// TIA Portal V20 export
Screen "PN_DIAGNOSTIC ETH P9P10"  1276x673
  ScreenItem "Line_Header_X0_Y64" at 0,64 size 1276x0  Type=HmiLine
  ScreenItem "Title_ScreenOverview_X390_Y2" at 390,2 size 500x30  Type=HmiTextBox
  ScreenItem "PN-Diag_Reset" at 93,2 size 90x60  Type=HmiButton
  ScreenItem "PN-Diag_ReadNew" at 184,2 size 90x60  Type=HmiButton
  ScreenItem "Textfeld_1" at 292,8 size 95x22  Type=HmiTextBox
  ScreenItem "LED_1_Left_2" at 0,0 size 100x30  Type=HmiCircle
  ScreenItem "LED_1_Left_1" at 0,0 size 100x30  Type=HmiCircle
  ScreenItem "Textfeld_4" at 292,35 size 95x22  Type=HmiTextBox
  ScreenItem "permanentareaborderrectangle" at 0,0 size 0x0  Type=HmiRectangle
  ScreenItem "Button_Back" at 2,2 size 90x60  Type=HmiButton
  ScreenItem "PN-Diag_Counters" at 1093,2 size 90x60  Type=HmiButton
  ScreenItem "PN-Diag_LegendᆉY2" at 1184,2 size 90x60  Type=HmiButton
  ScreenItem "Rectangle_1" at 51,92 size 203x123  Type=HmiRectangle
  ScreenItem "LSicar_DeviceDiag_7" at 485,101 size 170x97  Type=HmiFaceplateContainer
  ScreenItem "LSicar_DeviceDiag_2" at 292,273 size 171x97  Type=HmiFaceplateContainer
  ScreenItem "LSicar_DeviceDiag_4" at 81,101 size 170x97  Type=HmiFaceplateContainer
  ScreenItem "LSicar_DeviceDiag_11" at 293,101 size 170x105  Type=HmiFaceplateContainer
  ScreenItem "LSicar_DeviceDiag_3" at 1942,495 size 170x97  Type=HmiFaceplateContainer
  ScreenItem "LSicar_DeviceDiag_5" at 485,274 size 170x97  Type=HmiFaceplateContainer
  ScreenItem "LSicar_DeviceDiag_10" at 1604,81 size 170x97  Type=HmiFaceplateContainer
  ScreenItem "LSicar_DeviceDiag_6" at 2123,495 size 170x97  Type=HmiFaceplateContainer
  ScreenItem "LSicar_DeviceDiag_16" at 1375,728 size 170x97  Type=HmiFaceplateContainer
  ScreenItem "Faceplate container_1" at 880,104 size 170x100  Type=HmiFaceplateContainer
  ScreenItem "LSicar_DeviceDiag_13" at 2023,203 size 170x97  Type=HmiFaceplateContainer
  ScreenItem "线_4" at 190,162 size 60x0  Type=HmiLine
  ScreenItem "线_6" at 253,143 size 0x19  Type=HmiLine
  ScreenItem "线_26" at 254,142 size 129x0  Type=HmiLine
  ScreenItem "LSicar_DeviceDiag_17" at 61,269 size 170x105  Type=HmiFaceplateContainer
  ScreenItem "LSicar_DeviceDiag_18" at 680,101 size 170x97  Type=HmiFaceplateContainer
  ScreenItem "线_1" at 156,162 size 0x145  Type=HmiLine
  ScreenItem "线_3" at 363,152 size 23x0  Type=HmiLine
  ScreenItem "线_5" at 156,162 size 20x0  Type=HmiLine
  ScreenItem "线_7" at 363,153 size 0x54  Type=HmiLine
  ScreenItem "线_8" at 363,207 size 220x0  Type=HmiLine
  ScreenItem "线_9" at 583,179 size 0x27  Type=HmiLine
  ScreenItem "线_10" at 376,163 size 14x0  Type=HmiLine
  ScreenItem "线_11" at 376,163 size 0x54  Type=HmiLine
  ScreenItem "线_12" at 376,217 size 402x0  Type=HmiLine
  ScreenItem "线_13" at 778,179 size 0x37  Type=HmiLine
  ScreenItem "LSicar_DeviceDiag_20" at 1760,371 size 170x97  Type=HmiFaceplateContainer
  ScreenItem "LSicar_DeviceDiag_21" at 1941,371 size 170x97  Type=HmiFaceplateContainer
  ScreenItem "LSicar_DeviceDiag_22" at 2123,371 size 170x97  Type=HmiFaceplateContainer
  ScreenItem "LSicar_DeviceDiag_23" at 2309,371 size 170x97  Type=HmiFaceplateContainer
  ScreenItem "LSicar_DeviceDiag_24" at 1579,495 size 170x97  Type=HmiFaceplateContainer
  ScreenItem "LSicar_DeviceDiag_25" at 1760,495 size 170x97  Type=HmiFaceplateContainer
  ScreenItem "LSicar_DeviceDiag_26" at 1802,607 size 171x97  Type=HmiFaceplateContainer
  ScreenItem "Faceplate container_2" at 2309,495 size 170x97  Type=HmiFaceplateContainer
  ScreenItem "线_2" at 190,307 size 65x0  Type=HmiLine
  ScreenItem "线_14" at 255,307 size 0x81  Type=HmiLine
  ScreenItem "线_17" at 603,349 size 0x62  Type=HmiLine
  ScreenItem "线_24" at 255,389 size 157x0  Type=HmiLine
  ScreenItem "线_25" at 238,411 size 365x0  Type=HmiLine
  ScreenItem "线_15" at 412,349 size 0x40  Type=HmiLine
  ScreenItem "线_16" at 190,320 size 48x0  Type=HmiLine
  ScreenItem "线_18" at 238,320 size 0x90  Type=HmiLine
